(* IEC 61131-3 sources: Lasal-MCP/examples/SampleSource/2_PumpControlSolution/Stations/MachineControl/MachineControl/Class/SdiasSafetyManagerFSoE (part 2) *)

                          elsif (OptionalSettings.ModuleIDHBG = sHBG.usExpectedDeviceID) then
                            // the configured ID of LASAL and safety designer are equal

                            // if the module ID found is also the same => everthing is fine
                            if aModuleIDs[HBGPlace] = sHBG.usExpectedDeviceID then
                              MyPara.aPara[0] := _ClassOk$DINT;
                              CanActive := OldCanActive := TRUE;
                            else
                              // found something else
                              LogError("@02B4 (SdiasSafetyManagerFSoE::ClassSvr::NewInst) Wrong safety CAN terminal found (config of safety designer and hw classes match)");
                              MyPara.aPara[0] := _WrongHardware$DINT;
                              bHWConfigError := TRUE;
                            end_if;
                          else
                            // configuration of safety designer and hw classes does not match
                            LogError("@02B5 (SdiasSafetyManagerFSoE::ClassSvr::NewInst) Safety CAN terminal in hardware class configuration differs from safety designer configuration.");
                            MyPara.aPara[0] := _InvalidConfguration$DINT;
                            bHWConfigError := TRUE;
                          end_if;
                        else
                          MyPara.aPara[1] := SDIAS_SAFETY_INVALID_DEVICE_ID;

                          // projected in LASAL but not found in hardware
                          if sHBG.sdRequired then
                            MyPara.aPara[0] := _RequiredError$DINT;
                            bRequiredError := TRUE;
                            LogError("@02B6 (SdiasSafetyManagerFSoE::ClassSvr::NewInst) Required safety CAN terminal not available!");
                          else
                            // module is configured in safety designer
                            if (OptionalSettings.ModuleIDHBG <> SDIAS_SAFETY_INVALID_DEVICE_ID) then
                              // if the configuration does not match with the hardware classes
                              if (OptionalSettings.ModuleIDHBG <> sHBG.usExpectedDeviceID) then
                                LogError("@02B5 (SdiasSafetyManagerFSoE::ClassSvr::NewInst) Safety CAN terminal in hardware class configuration differs from safety designer configuration.");
                                MyPara.aPara[0] := _InvalidConfguration$DINT;
                                bHWConfigError := TRUE;

                              // the IDs match but it's not optional. since it's not available => error
                              elsif (OptionalSettings.OptionalFlagHBG.1 = FALSE) then
                                MyPara.aPara[0] := _NoHardware$DINT;
                                LogError("@02B7 (SdiasSafetyManagerFSoE::ClassSvr::NewInst) Could not find the non-optional Safety CAN terminal defined in the safety designer configuration.");
                                bHWConfigError := TRUE;

                              else
                                // if the IDs match and it's optional => just show no hardware (no error)
                                MyPara.aPara[0] := _NoHardware$DINT;
                              end_if;
                            else
                              LogError("@02B8 (SdiasSafetyManagerFSoE::ClassSvr::NewInst) Safety CAN terminal in hardware class configuration but not physically available and not in safety designer configuration.");
                              MyPara.aPara[0] := _NoHardware$DINT;
                            end_if;
                          end_if;
                        end_if;
                        sHBG.pThis^.NewInst(#MyPara, #MyResult);
                      else
                        // nothing projected for HBG in the lasal project

                        // if module is configured in safety designer
                        if (OptionalSettings.ModuleIDHBG <> SDIAS_SAFETY_INVALID_DEVICE_ID) then
                          // if a HBG has been found
                          if HBGPlace <> SDIAS_SAFETY_INVALID_MAX_PLACE then
                            // if it's not the configured module
                            if (aModuleIDs[HBGPlace] <> OptionalSettings.ModuleIDHBG) then
                              LogError("@02B9 (SdiasSafetyManagerFSoE::ClassSvr::NewInst) Safety CAN terminal found doesn't match the safety designer configuration.");
                              bHWConfigError := TRUE;
                            end_if;
                          else
                            // module not available (only a problem if it's not optional)
                            if (OptionalSettings.OptionalFlagHBG.1 = FALSE) then
                              LogError("@02BA (SdiasSafetyManagerFSoE::ClassSvr::NewInst) Could not find the non-optional Safety CAN terminal defined in the safety designer configuration.");
                              bHWConfigError := TRUE;
                            end_if;
                          end_if;
                        else
                          // module not configured in safety designer. if there is a module available, the number of IOs in safety does not match the config
                          if HBGPlace <> SDIAS_SAFETY_INVALID_MAX_PLACE then
                            LogError("@02BB (SdiasSafetyManagerFSoE::ClassSvr::NewInst) Safety CAN terminal found but not projected in the safety designer configuration.");
                            bHWConfigError := TRUE;
                          end_if;
                        end_if;
                      end_if;
                    else
                      // old firmware (no optional settings available)
                      if MaxPlace <> SDIAS_SAFETY_INVALID_MAX_PLACE then
                        pSafetyModuleInfo := #aSafetyModuleInfo[0];

                        // always the same command
                        MyPara.uiCmd := SDIAS_SET_CLASS_STATE;

                        for i := 0 to MaxPlace do
                          if pSafetyModuleInfo^.pThis then
                            MyPara.aPara[1] := aModuleIDs[i];
                            if aModuleIDs[i] = pSafetyModuleInfo^.usExpectedDeviceID then
                              MyPara.aPara[0] := _ClassOk$DINT;
                            elsif aModuleIDs[i] <> SDIAS_SAFETY_INVALID_DEVICE_ID then
                              if pSafetyModuleInfo^.sdRequired then
                                MyPara.aPara[0] := _RequiredError$DINT;
                                bRequiredError := TRUE;
                                LogValue("@02AC (SdiasSafetyManagerFSoE::ClassSvr::NewInst) Wrong safety IO module at required place {0}.", Value:=i);
                              else
                                MyPara.aPara[0] := _WrongHardware$DINT;
                                bHWConfigError  := TRUE;
                              end_if;
                            else
                              if pSafetyModuleInfo^.sdRequired then
                                MyPara.aPara[0] := _RequiredError$DINT;
                                bRequiredError := TRUE;
                                LogValue("@02AB (SdiasSafetyManagerFSoE::ClassSvr::NewInst) No safety IO module at required place {0}.", Value:=i);
                              else
                                MyPara.aPara[0] := _NoHardware$DINT;
                                // Hardwareclass placed in Project but no physical Hardware available is allowed
                                // bHWConfigError  := TRUE;
                              end_if;
                            end_if;
                            pSafetyModuleInfo^.pThis^.NewInst(#MyPara, #MyResult);

                          elsif aModuleIDs[i] <> SDIAS_SAFETY_INVALID_DEVICE_ID then  // HWK this pointer is NIL but a module is identified
                            bHWConfigError  := TRUE;
                          end_if;

                          pSafetyModuleInfo += sizeof(t_SdiasSafetyModuleInfo);
                        end_for;
                      end_if;

                      // Check if a module info was passed for which there is no corrosponding HWK object.
                      if MaxPlace + 1 < sizeof(t_ModuleIDs) then
                        // it's only a config error if it's not the HBG
                        if (aModuleIDs[MaxPlace + 1] <> SDIAS_SAFETY_INVALID_DEVICE_ID) & ((MaxPlace + 1) <> HBGPlace) then
                          bHWConfigError  := TRUE;
                        end_if;
                      end_if;

                      // check for hbg
                      if sHBG.pThis then
                        MyPara.uiCmd := SDIAS_SET_CLASS_STATE;
                        if HBGPlace <> SDIAS_SAFETY_INVALID_MAX_PLACE then
                          MyPara.aPara[1] := aModuleIDs[HBGPlace];

                          if aModuleIDs[HBGPlace] = sHBG.usExpectedDeviceID then
                            MyPara.aPara[0] := _ClassOk$DINT;
                            CanActive := OldCanActive := TRUE;
                            bHWConfigError := FALSE;
                          elsif aModuleIDs[HBGPlace] <> SDIAS_SAFETY_INVALID_DEVICE_ID then
                            if sHBG.sdRequired then
                              MyPara.aPara[0] := _RequiredError$DINT;
                              bRequiredError := TRUE;
                              LogError("@02BE (SdiasSafetyManagerFSoE::ClassSvr::NewInst) Wrong safety IO module at required HBG place.");
                            else
                              MyPara.aPara[0] := _WrongHardware$DINT;
                              CanActive := OldCanActive := FALSE;
                            end_if;
                          else
                            if sHBG.sdRequired then
                              MyPara.aPara[0] := _RequiredError$DINT;
                              bRequiredError := TRUE;
                              LogError("@02BF (SdiasSafetyManagerFSoE::ClassSvr::NewInst) HBG required but not available!");
                            else
                              MyPara.aPara[0] := _NoHardware$DINT;
                              CanActive := OldCanActive := FALSE;
                            end_if;
                          end_if;
                        else
                          MyPara.aPara[1] := SDIAS_SAFETY_INVALID_DEVICE_ID;
                          if sHBG.sdRequired then
                            MyPara.aPara[0] := _RequiredError$DINT;
                            bRequiredError := TRUE;
                            LogError("@02BE (SdiasSafetyManagerFSoE::ClassSvr::NewInst) Wrong safety IO module at required HBG place.");
                          else
                            MyPara.aPara[0] := _WrongHardware$DINT;
                            CanActive := OldCanActive := FALSE;
                          end_if;
                        end_if;
                        sHBG.pThis^.NewInst(#MyPara, #MyResult);
                      end_if;
                    end_if;

                    if bRequiredError then
                      MyPara.uiCmd := _BUS_IF_SET_REQUIRED_ERROR;
                      ToBusInterface.NewInst(#MyPara, #MyResult);
                    end_if;

                    if bHWConfigError then
                      // if we have optional settings, we already logged the reason
                      if b_GotOptionalSettings = FALSE then
                        LogError("@ß02C0 (SdiasSafetyManagerFSoE::ClassSvr::NewInst) Hardwareconfiguration does not match objects placed in network.");
                      end_if;

                      // Check if Safetymanyger is required
                      MyPara.uiCmd     := _BUS_IF_GET_REQUIRED_SETTING;
                      ToBusInterface.NewInst(pPara:=#MyPara, pResult:=#MyResult);
                      if MyResult.aData[0]$t_BusIFRetvalErrorcode = _BUS_IF_RETVAL_OK then
                        // if it's required => set required error
                        if MyResult.aData[4] then

                          MyPara.uiCmd := _BUS_IF_SET_REQUIRED_ERROR;
                          ToBusInterface.NewInst(#MyPara, #MyResult);
                        else

                          SetSafetyState(_WrongSafetyHW);
                          Online      := 0;

                          // Update BusIF ClassState
                          MyPara.uiCmd := _BUS_IF_SET_CLASS_STATE;
                          MyPara.aPara[0] := _WrongHardware$DINT;
                          ToBusInterface.NewInst(#MyPara, #MyResult);

                          // Cancel init
                          eInitSSWErrorStep := eInitSSW;
                          eInitSSW := _InitError;

                          // Set Module states
                          pSafetyModuleInfo := #aSafetyModuleInfo[0];
                          // always the same command
                          MyPara.uiCmd := SDIAS_SET_CLASS_STATE;
                          MyPara.aPara[0] := _ModuleFoundButManagerIsOff$DINT;

                          if MaxPlace <> SDIAS_SAFETY_INVALID_MAX_PLACE then
                            for i := 0 to MaxPlace do
                              if pSafetyModuleInfo^.pThis then
                                MyPara.aPara[1] := aModuleIDs[i];
                                pSafetyModuleInfo^.pThis^.NewInst(#MyPara, #MyResult);
                              end_if;
                              pSafetyModuleInfo += sizeof(t_SdiasSafetyModuleInfo);
                            end_for;
                          end_if;

                          // check for hbg
                          if sHBG.pThis then
                            sHBG.pThis^.NewInst(#MyPara, #MyResult);
                          end_if;

                        end_if;

                      end_if;

                    end_if;

                  else
                    LogError("@02C1 (SdiasSafetyManagerFSoE::ClassSvr::NewInst) Invalid SDO response buffer pointer.");
                  end_if;
                else
                  LogError("@02C2 (SdiasSafetyManagerFSoE::ClassSvr::NewInst) Invalid length for SDO response data.");
                end_if;

                eResponseState := _valid;
              else
                LogError("@02C3 (SdiasSafetyManagerFSoE::ClassSvr::NewInst) SDO response arrived when no response was expected.");
              end_if;
            end_if;
          elsif (LastSDO.Command = _BUS_IF_READ_VIA_SDO_CTRL) then
            if LastSDO.ResponseArrived = FALSE then
              if pPara^.aPara[5] = LastSDO.Length then
                if pPara^.aPara[4] then
                  // all parameters are fine, so we're ready
                  ret_code := READY;

                  // copy the response data
                  _memcpy(ptr1:=Config.pActData, ptr2:=pPara^.aPara[4]$pVoid, cntr:=LastSDO.Length);
                else
                  LogError("@02C1 (SdiasSafetyManagerFSoE::ClassState::NewInst) Invalid SDO response buffer pointer.");
                end_if;
              else
                LogError("@02C2 (SdiasSafetyManagerFSoE::ClassState::NewInst) Invalid length for SDO response data.");
              end_if;

              LastSDO.ResponseArrived := TRUE;
            else
              LogError("@02C3 (SdiasSafetyManagerFSoE::ClassState::NewInst) SDO response arrived when no response was expected.");
            end_if;
          elsif (LastSDO.Command = _BUS_IF_WRITE_VIA_SDO_CTRL) then
            if LastSDO.ResponseArrived = FALSE then
              // all parameters are fine, so we're ready
              ret_code := READY;

              LastSDO.ResponseArrived := TRUE;
            else
              LogError("@02C3 (SdiasSafetyManagerFSoE::ClassState::NewInst) SDO response arrived when no response was expected.");
            end_if;
          end_if;
        else
          LogError("@02C4 (SdiasSafetyManagerFSoE::ClassSvr::NewInst) SDO transfer failed.");
        end_if;
      else
        LogError("@02C5 (SdiasSafetyManagerFSoE::ClassSvr::NewInst) Received invalid SDO response.");
      end_if;

//**********************************************************************************************************************************************************
    _BUS_IF_DATA_POINTER_AVAILABLE:
      // does nothing in the FSoE version
      ret_code := READY;

//**********************************************************************************************************************************************************
    _BUS_IF_RESET_DETECTED:
      // don't overwrite other errors
      if SafetyState = _SafetyClassOK then
        SafetyState := _LostPowerSupply;
      end_if;

      // check if module is requred
      MyPara.uiCmd     := _BUS_IF_GET_REQUIRED_SETTING;
      ToBusInterface.NewInst(pPara:=#MyPara, pResult:=#MyResult);
      if MyResult.aData[0]$t_BusIFRetvalErrorcode = _BUS_IF_RETVAL_OK then
        // if it's required => set required error
        if MyResult.aData[4] then

          MyPara.uiCmd := _BUS_IF_SET_REQUIRED_ERROR;
          ToBusInterface.NewInst(#MyPara, #MyResult);
        end_if;
      end_if;

      // drop config of connected modules

      // initialize the message for the periphery
      MyPara.uiCmd := SDIAS_SET_CLASS_STATE;
      MyPara.aPara[1] := 0;// no device ID
      MyPara.aPara[0] := _NoHardware$DINT;

      // tell the connected IO module objects
      if MaxPlace <> SDIAS_SAFETY_INVALID_MAX_PLACE then
        pSafetyModuleInfo := #aSafetyModuleInfo[0];

        for i := 0 to MaxPlace do
          if pSafetyModuleInfo^.pThis then
            pSafetyModuleInfo^.pThis^.NewInst(#MyPara, #MyResult);
          end_if;

          pSafetyModuleInfo += sizeof(t_SdiasSafetyModuleInfo);
        end_for;
      end_if;

      // tell the hbg (if available)
      if sHBG.pThis then
        sHBG.pThis^.NewInst(#MyPara, #MyResult);
      end_if;

//**********************************************************************************************************************************************************
    _BUS_IF_RESET_GONE_DETECTED:
      if SafetyState = _LostPowerSupply then

        // get safety and serial numbers of connected modules
        bUpdateModuleConfig := TRUE;

        // remember the time. in case we don't get the SDO response to signal the firmware being ready, we use a timeout
        ud_ResetGoneTime := ops.tAbsolute;

        // we wait for an asynchronous SDO response in the cyclic of the base class. once we got that, the firmware is ready
        b_WaitForFirmwareBoot := TRUE;

        // refetch IDs of connected modules
        eCheckIDSSW := _Wait4Idle;

        SafetyState := _SafetyClassOK;
      end_if;

//**********************************************************************************************************************************************************

    CMD_GET_HARDWARE_DIAGNOSIS:
      //Returns module info
      ret_code := ERROR;
      pResult^.aData[0]$t_HWCGetHardwareDiagnosisOut.retcode := _HWC_RETVAL_ERROR;

      pStr_HWTRequested := pPara^.aPara[0]$t_HWCGetHardwareDiagnosisIn.pStr_HardewareTreeEntry;

      tmpplace := (pStr_HWTRequested+pPara^.aPara[0]$t_HWCGetHardwareDiagnosisIn.us_current_index)^$USINT;

      //Check if pointer is valid
      if aSafetyModuleInfo[tmpplace].pThis then

        // Set Offline Device ID
        pResult^.aData[0]$t_HWCGetHardwareDiagnosisOut.ud_DeviceID := (aSafetyModuleInfo[tmpplace].usExpectedDeviceID AND 2#00111000 ) shr 3;   // Bit 3-5 Modul typ
        pResult^.aData[0]$t_HWCGetHardwareDiagnosisOut.ud_Variante :=  aSafetyModuleInfo[tmpplace].usExpectedDeviceID AND 2#00000111;  // Bit 0-2 Submodul typ

        if aModuleIDs[tmpplace] = aSafetyModuleInfo[tmpplace].usExpectedDeviceID then

          ret_code := READY;
          pResult^.aData$t_HWCGetHardwareDiagnosisOut.retcode := _HWC_RETVAL_OK;

          pResult^.aData[0]$t_HWCGetHardwareDiagnosisOut.ud_DeviceID  := (aModuleIDs[tmpplace] AND 2#00111000 ) shr 3;  // Bit 3-5 Modul typ
          pResult^.aData[0]$t_HWCGetHardwareDiagnosisOut.ud_Variante  :=  aModuleIDs[tmpplace] AND 2#00000111; // // Bit 0-2 Submodul typ
          pResult^.aData[0]$t_HWCGetHardwareDiagnosisOut.ud_Place     := tmpplace;

          // Get Serialno ---------------------------------------------------------------------------------------------
          _memcpy(ptr1 := #a_SerialNo[0]
                , ptr2 := #sSafetySerNrs.aSerialNumbers[tmpplace]
                , cntr := sizeof(sSafetySerNrs.aSerialNumbers[tmpplace]) );

          a_SerialNo[sizeof(sSafetySerNrs.aSerialNumbers[tmpplace])] := 0;  // 0 Terminierung

          pResult^.aData[0]$t_HWCGetHardwareDiagnosisOut.pStr_SerialNo := #a_SerialNo[0];

          pResult^.aData[0]$t_HWCGetHardwareDiagnosisOut.hd_SafetyNumber  := sSafetySerNrs.aSafetyNumbers[tmpplace];

          // first free the old then create the memory (linked list) for the additional information

          if pAdditionalDiagInfo then
            HwDiagFreeDynExtList(pList:=pAdditionalDiagInfo);
          end_if;
          pAdditionalDiagInfo      := NIL;

          // add the firmware version
          pNewElement := HwDiagAddDynExt2List(ppList:=#pAdditionalDiagInfo, EntryID:=_HWC_DIAG_ID_SAFETY_FIRMWARE_VERSION, udVersion:=1, udDataLength:=sizeof(HDINT));

          if pNewElement then
            // add the data in the reserved memory
            (pNewElement$^HDINT + sizeof(t_HWCGetHardwareDiagnosisOutDynExt))^ := FirmwareVersion;
          end_if;

          // add the safety designer project name
          pNewElement := HwDiagAddDynExt2List(ppList:=#pAdditionalDiagInfo, EntryID:=_HWC_DIAG_ID_SAFETY_DESIGNER_PROJECT_NAME, udVersion:=1, udDataLength:=ProjectNameStr.GetLength());

          if pNewElement then
            // add the data in the reserved memory
            ProjectNameStr.ReadDataOff(udOff:=0, pData:=pNewElement$^USINT + sizeof(t_HWCGetHardwareDiagnosisOutDynExt), udMax:=pNewElement^.ud_DataLength);
          end_if;

          // add the safety designer project revision
          pNewElement := HwDiagAddDynExt2List(ppList:=#pAdditionalDiagInfo, EntryID:=_HWC_DIAG_ID_SAFETY_DESIGNER_PROJECT_REVISION, udVersion:=1, udDataLength:=ProjectRevisionStr.GetLength());

          if pNewElement then
            // add the data in the reserved memory
            ProjectRevisionStr.ReadDataOff(udOff:=0, pData:=pNewElement$^USINT + sizeof(t_HWCGetHardwareDiagnosisOutDynExt), udMax:=pNewElement^.ud_DataLength);
          end_if;

          pResult^.aData[0]$t_HWCGetHardwareDiagnosisOut.p_DynExtList := pAdditionalDiagInfo;

        elsif aModuleIDs[tmpplace] <> SDIAS_SAFETY_INVALID_DEVICE_ID then
          pResult^.aData$t_HWCGetHardwareDiagnosisOut.retcode := _HWC_RETVAL_ERROR_WRONG_HARDWARE;
        else
          pResult^.aData$t_HWCGetHardwareDiagnosisOut.retcode := _HWC_RETVAL_ERROR_NO_HARDWARE;
        end_if;

      else
        pResult^.aData[0]$t_HWCGetHardwareDiagnosisOut.retcode := _HWC_RETVAL_ERROR_SDIAS_MODULE_NOT_FOUND;
      end_if;

//**********************************************************************************************************************************************************
    CMD_GET_HARDWARE_TREE_ENTRY:
      //Returns module info

      ret_code := ERROR;
      pResult^.aData[0]$t_HWCGetHardwareTreeEntryOut.retcode := _HWC_RETVAL_ERROR;

      pStr_HWTreeEntry := pPara^.aPara[0]$t_HWCGetHardwareTreeEntryIn.pStr_LastHardewareTreeEntry;

      //First HWT Path
      if (pStr_HWTreeEntry + pStr_HWTreeEntry$^UINT^)^ <> HWT_ESCAPE_INTERNALBUS_SDIAS_SAFETY then  // + 1 for Byte length -1 for 2nd last element of string

        if aSafetyModuleInfo[0].pThis then

          _memcpy(ptr1 := #a_HWTEntryStr[0]
                , ptr2 := pPara^.aPara[0]$t_HWCGetHardwareTreeEntryIn.pStr_LastHardewareTreeEntry
                , cntr := pPara^.aPara[0]$t_HWCGetHardwareTreeEntryIn.pStr_LastHardewareTreeEntry$^UINT^ +2 );  // +2 2 Byte Strlength is not included in the stringlength

          // Add escape sequence
          a_HWTEntryStr[0]$UINT += 1;
          a_HWTEntryStr[a_HWTEntryStr[0]$UINT+1] := HWT_ESCAPE_INTERNALBUS_SDIAS_SAFETY;

          // Add Place
          a_HWTEntryStr[0]$UINT += 1;
          a_HWTEntryStr[a_HWTEntryStr[0]$UINT+1] := 0;

          //Return Hardware Tree Entry and set return codes
          pResult^.aData[0]$t_HWCGetHardwareTreeEntryOut.pStr_NextHardewareTreeEntry := #a_HWTEntryStr[0];

          pResult^.aData[0]$t_HWCGetHardwareTreeEntryOut.retcode := _HWC_RETVAL_OK_HWTSTR_RETURNED;
          ret_code := READY;

        else
          pResult^.aData[0]$t_HWCGetHardwareTreeEntryOut.retcode := _HWC_RETVAL_ERROR_SDIAS_MODULE_NOT_FOUND;
        end_if;

      //search next module
      else

        usNextPlace := (pStr_HWTreeEntry  + pPara^.aPara[0]$t_HWCGetHardwareTreeEntryIn.us_current_index)^$USINT+1;

        if usNextPlace <= SDIAS_SAFETY_MAX_PLACE_NR &
           aSafetyModuleInfo[usNextPlace].pThis then

          _memcpy(ptr1 := #a_HWTEntryStr[0]
                , ptr2 := pPara^.aPara[0]$t_HWCGetHardwareTreeEntryIn.pStr_LastHardewareTreeEntry
                , cntr := pPara^.aPara[0]$t_HWCGetHardwareTreeEntryIn.pStr_LastHardewareTreeEntry$^UINT^ +2 );  // +2 2 Byte Strlength is not included in the stringlength

          // Set new Place
          a_HWTEntryStr[a_HWTEntryStr[0]$UINT + 1] := usNextPlace;

          pResult^.aData[0]$t_HWCGetHardwareTreeEntryOut.pStr_NextHardewareTreeEntry := #a_HWTEntryStr[0];

          //Return Hardware Tree Entry and set return codes
          pResult^.aData[0]$t_HWCGetHardwareTreeEntryOut.retcode := _HWC_RETVAL_OK_HWTSTR_RETURNED;
          ret_code := READY;

        else
          ret_code := READY;
          pResult^.aData$t_HWCGetHardwareTreeEntryOut.retcode := _HWC_RETVAL_OK_END_OF_LIST;
        end_if;
      end_if;

//**********************************************************************************************************************************************************

//*****************************************************************************
//** INTERNAL COMMANDS                                                       **
//*****************************************************************************

//**********************************************************************************************************************************************************
    CMD_SM_READ_PDO_SIZE:
      // get the size of the PDO
      LastSDO.Command := _BUS_IF_READ_VIA_SDO;
      LastSDO.Offset  := SBF_OFFSET_SPDO_LENGTH;
      LastSDO.Length  := sizeof(UINT);

      MyPara.uiCmd    := LastSDO.Command$UINT;
      MyPara.aPara[0] := LastSDO.Offset;
      MyPara.aPara[1] := LastSDO.Length;
      ret_code := ToBusInterface.NewInst(#MyPara, #MyResult);

//**********************************************************************************************************************************************************
  else
    ret_code := SafetyBaseFSoE::NewInst(pPara, pResult);
//**********************************************************************************************************************************************************
  END_CASE;

END_FUNCTION

FUNCTION VIRTUAL SdiasSafetyManagerFSoE::ShowProjectRevision

  ProjectNameStr.WriteDataOff(udLen:=PrjNameStrLen + 1, udOff:=0, pData:=pPrjNameStr);

  ProjectRevisionStr.WriteDataOff(udLen:=PrjRevStrLen + 1, udOff:=0, pData:=pPrjRevStr);

END_FUNCTION

FUNCTION VIRTUAL SdiasSafetyManagerFSoE::InitSafeModule
  VAR_OUTPUT
    sd_retval 	: DINT;
  END_VAR

  // allocate memory for finding unsafe-IO-Servers
  // in first place we allocate 512 byte for our blocked transfers
  p_BlockedTransferMemory := ToStdLib.Malloc( size := SBF_CONFIG_MEMORY_BLOCK_SIZE );
  IF p_BlockedTransferMemory <> NIL THEN
    ud_BlockedTransferMemorySize := SBF_CONFIG_MEMORY_BLOCK_SIZE;
  ELSE
    SafetyState := _MemAllocFailed;
    sd_retval := -100;
    return;
  END_IF;

  // if there is a safety manager to gather the configuration
  if pSafetyManagerThis then
    // allocate memory for gathering configuration information => in first place we allocate 512 byte
    pConfigMem := ToStdLib.Malloc( size := SBF_CONFIG_MEMORY_BLOCK_SIZE );
    IF pConfigMem <> NIL THEN
      ConfigMemSize := SBF_CONFIG_MEMORY_BLOCK_SIZE;
      ConfigMemSizeUsed := 4;
    ELSE
      SafetyState := _MemAllocFailed;
      sd_retval := -100;
      return;
    END_IF;
  end_if;

END_FUNCTION

FUNCTION VIRTUAL GLOBAL SdiasSafetyManagerFSoE::CanOut::NewInst
  VAR_INPUT
    pPara 	: ^CmdStruct;
    pResult 	: ^results;
  END_VAR
  VAR_OUTPUT
    ret_code 	: iprStates;
  END_VAR
  VAR
    tempCmd         : CmdStruct;
    _result         : results;
  END_VAR

  CASE pPara^.uiCmd OF
//**********************************************************************************************************************************************************
    SDIAS_SAFETY_LOGIN_HBG:
      // check parameters
      if pPara^.aPara[0] & pPara^.aPara[1] then

        sHBG.pThis               := pPara^.aPara[0]$pVirtualBase;
        sHBG.usExpectedDeviceID  := pPara^.aPara[1]$USINT;
        sHBG.sdRequired          := pPara^.aPara[2];
        sHBG.pIOStates           := pPara^.aPara[3]$^HDINT;

        // if leds/hgb not added so far, add them
        if StateBytesUsed = 0 then
          StateBitsUsed := (sizeof(t_LedAndIOStates.biLEDs) + sizeof(t_LedAndIOStates.HBGInputs)) * 8;
          // refresh state bytes used value
          StateBytesUsed := ((StateBitsUsed-1) / 8) + 1;
        end_if;

        if sHBG.sdRequired & (b_AnyModuleRequired = FALSE) then
          b_AnyModuleRequired := TRUE;
          // if any access is required => the businterface is also required
          tempCmd.uiCmd := _BUS_IF_SET_REQUIRED;
          ToBusInterface.NewInst(pPara:=#tempCmd, pResult:=#_result);
          if _result.aData[0]$t_BusIFRetvalErrorcode <> _BUS_IF_RETVAL_OK then
            LogError("@029D (SdiasSafetyManagerFSoE::CanOut::NewInst) Failed to set the BusInterface to required.");
          end_if;
        end_if;
      else
        ret_code := ERROR;
      end_if;
//**********************************************************************************************************************************************************
  END_CASE;

  ret_code := READY;

END_FUNCTION

FUNCTION VIRTUAL SdiasSafetyManagerFSoE::GetConfiguration
  VAR
    pHelp                 : ^void;
    SizeToGo              : UINT;
    ActSize               : UINT;
    ActAddr               : HDINT;
    SDOReqBuf             : SDORequReadConfig;
    SDORspBuf             : ARRAY [0..SBF_SDO_MAX_LENGTH-1] OF USINT;
    pRspBuf               : ^SDORespReadConfig;
    i                     : DINT;
    pSafetyModuleInfo     : ^t_SdiasSafetyModuleInfo;
    MyPara 	              : CmdStruct;
    MyResult              : Results;
  END_VAR

  //initialize header-data for request

  //calculate length without crc
  SDOReqBuf.StdHeader.Len := sizeof(SDORequReadConfig) - sizeof(SDOHeader.StdHeader.CRC);

  //type
  SDOReqBuf.StdHeader.Typ := SDO_STD;

  //command for reading config data
  SDOReqBuf.StdHeader.Cmd := SBF_SDO_COMMAND_READ;

  // read the complete 256 Bytes of safety and serial number info
  pHelp    := #sSafetySerNrs;
  SizeToGo := sizeof(sSafetySerNrs);
  pRspBuf  := (#SDORspBuf)$^SDORespReadConfig;
  ActAddr  := SBF_SDO_ADDRESS_SER_NR_DATA;

  while SizeToGo do
    if SizeToGo > SDIAS_SAFTEY_SDO_MAX_DATA_PER_PAKET then
      ActSize := SDIAS_SAFTEY_SDO_MAX_DATA_PER_PAKET;
    else
      ActSize := SizeToGo;
    end_if;

    if SDOReadCfgRequ(p_SDORequestBuffer  := #SDOReqBuf,
                      p_SDOResponseBuffer := pRspBuf,
                      ud_Address          := ActAddr,
                      us_Length           := ActSize$USINT,
                      b_UseCache          := FALSE) then
      LogError("@02C6 (SdiasSafetyManagerFSoE::GetConfiguration) Failed to get safety and serial numbers of the IO modules.");
      return;
    else
      _memcpy(ptr1:=pHelp, ptr2:=#pRspBuf^.ud_Data, cntr:=ActSize);
    end_if;

    SizeToGo  -= ActSize;
    ActAddr   += ActSize;
    pHelp     += ActSize;
  end_while;

  // read the complete 64 Bytes of hardware version info
  pHelp    := #sHwVersions;
  SizeToGo := sizeof(sHwVersions);
  pRspBuf  := (#SDORspBuf)$^SDORespReadConfig;
  ActAddr  := SBF_SDO_ADDRESS_HW_VERSIONS;

  while SizeToGo do
    if SizeToGo > SDIAS_SAFTEY_SDO_MAX_DATA_PER_PAKET then
      ActSize := SDIAS_SAFTEY_SDO_MAX_DATA_PER_PAKET;
    else
      ActSize := SizeToGo;
    end_if;

    if SDOReadCfgRequ(p_SDORequestBuffer  := #SDOReqBuf,
                      p_SDOResponseBuffer := pRspBuf,
                      ud_Address          := ActAddr,
                      us_Length           := ActSize$USINT,
                      b_UseCache          := FALSE) then
      LogError("@02F9 (SdiasSafetyManagerFSoE::GetConfiguration) Failed to get hw versions of the Safe IO modules!");
      return;
    else
      // if the return code in the response buffer is not 0 => the virtual memory is not available
      if pRspBuf^.us_Returncode <> 0 then
        // reset array to make sure there are no hw versions stored
        _memset(dest:=#sHwVersions.aVersion[0], usByte:=0, cntr:=sizeof(sHwVersions));
        exit;
      end_if;

      _memcpy(ptr1:=pHelp, ptr2:=#pRspBuf^.ud_Data, cntr:=ActSize);
    end_if;

    SizeToGo  -= ActSize;
    ActAddr   += ActSize;
    pHelp     += ActSize;
  end_while;

  // only available for IOs, not the HBG
  if MaxPlace <> SDIAS_SAFETY_INVALID_MAX_PLACE then
    // always the same command
    MyPara.uiCmd := SDIAS_SET_NUMBERS;

    pSafetyModuleInfo := #aSafetyModuleInfo[0];
    for i := 0 to MaxPlace$DINT do
      // safety number
      MyPara.aPara[0] := (sSafetySerNrs.aSafetyNumbers[i])$DINT;

      // pointer to serial number string
      MyPara.aPara[1] := (#sSafetySerNrs.aSerialNumbers[i][0])$DINT;

      // hw version
      MyPara.aPara[2] := (sHwVersions.aVersion[i])$DINT;

      pSafetyModuleInfo^.pThis^.NewInst(#MyPara, #MyResult);

      pSafetyModuleInfo += sizeof(t_SdiasSafetyModuleInfo);
    end_for;
  end_if;

END_FUNCTION

FUNCTION VIRTUAL GLOBAL SdiasSafetyManagerFSoE::DisconnectEvent
  VAR
    i                 : UDINT;
    pSafetyModuleInfo : ^t_SdiasSafetyModuleInfo;
    MyPara 	          : CmdStruct;
    MyResult          : Results;
  END_VAR

  SafetyBaseFSoE::DisconnectEvent();

  // initialize the message for the periphery
  MyPara.uiCmd := SDIAS_SET_CLASS_STATE;
  MyPara.aPara[1] := 0;// no device ID
  MyPara.aPara[0] := _NoHardware$DINT;

  // tell the connected IO module objects
  if MaxPlace <> SDIAS_SAFETY_INVALID_MAX_PLACE then
    pSafetyModuleInfo := #aSafetyModuleInfo[0];

    for i := 0 to MaxPlace do
      if pSafetyModuleInfo^.pThis then
        pSafetyModuleInfo^.pThis^.NewInst(#MyPara, #MyResult);
      end_if;

      pSafetyModuleInfo += sizeof(t_SdiasSafetyModuleInfo);
    end_for;
  end_if;

  // tell the hbg (if available)
  if sHBG.pThis then
    sHBG.pThis^.NewInst(#MyPara, #MyResult);
  end_if;

  // clear the strings
  ProjectNameStr.Clear();
  ProjectRevisionStr.Clear();

END_FUNCTION

FUNCTION VIRTUAL SdiasSafetyManagerFSoE::SetSafetyState
  VAR_INPUT
    NewState 	: SafetyConfigStateType;
  END_VAR
  VAR
    MyPara 	  : CmdStruct;
    MyResult	: results;
  END_VAR

  // use it locally
  SafetyState := NewState;

  // tell the outer class
  MyPara.uiCmd := SDIAS_SET_SAFETY_STATE;
  MyPara.aPara[0] := NewState$DINT;
  ToBusInterface.NewInst(#MyPara, #MyResult);

END_FUNCTION

FUNCTION VIRTUAL GLOBAL SdiasSafetyManagerFSoE::CyWork
  VAR_INPUT
    EAX 	: UDINT;
  END_VAR
  VAR_OUTPUT
    state (EAX) 	: UDINT;
  END_VAR
  VAR
    MyPara 	          : CmdStruct;
    MyResult          : Results;
    TmpRetCode        : iprStates;
  END_VAR

  // if the initialisiation has been finished and there is an object for the hbg check if it's has been connected or disconnected
  if Online then

    case eCheckIDSSW of
  //**********************************************************************************************************************************************************
      _Nothing:
        if sHBG.pThis then
          // check for a can connect event
          if CanActive > OldCanActive then
            // if we're already idle => get it on
            if eResponseState = _idle then
              eCheckIDSSW := _GetIDs;
            else
              // otherwise, wait for it (need to remember the connect event)
              eCheckIDSSW := _Wait4Idle;
            end_if;

          // check for a can disconnect event
          elsif CanActive < OldCanActive then
            if sHBG.sdRequired then
              // if it's required => required error
              MyPara.uiCmd := _BUS_IF_SET_REQUIRED_ERROR;
              ToBusInterface.NewInst(#MyPara, #MyResult);
            else
              // otherwise show that it has been disconnected
              MyPara.uiCmd := SDIAS_SET_CLASS_STATE;
              MyPara.aPara[1] := 0;// no device ID
              MyPara.aPara[0] := _NoHardware$DINT;
              sHBG.pThis^.NewInst(#MyPara, #MyResult);
            end_if;
          end_if;
          OldCanActive := CanActive;
        end_if;

  //**********************************************************************************************************************************************************
      _Wait4Idle:
        if eResponseState = _idle then
          eCheckIDSSW := _GetIDs;
        end_if;

  //**********************************************************************************************************************************************************
      _GetIDs:
        case eResponseState of
        //*****************************************************
          _idle:
            LastSDO.Command := _BUS_IF_READ_VIA_SDO;
            LastSDO.Offset  := SBF_OFFSET_IO_MODULE_IDS;
            LastSDO.Length  := sizeof(t_ModuleIDs);

            MyPara.uiCmd    := LastSDO.Command$UINT;
            MyPara.aPara[0] := LastSDO.Offset;
            MyPara.aPara[1] := LastSDO.Length;
            TmpRetcode := ToBusInterface.NewInst(#MyPara, #MyResult);
            if TmpRetcode = READY then
              SDOTimeMark  := ops.tAbsolute;
              eResponseState:= _wait;
            elsif TmpRetcode = ERROR then
              LogError("@02A7 (SdiasSafetyManagerFSoE::InitModule) Failed to add read SDO for module configuration.");
            end_if;
        //*****************************************************
          _wait:
            // wait for response
            if ((ops.tAbsolute - SDOTimeMark) > SDIAS_SAFTEY_SDO_RESPONSE_TIMEOUT) then
              LogError("@02A1 (SdiasSafetyManagerFSoE::InitModule) SDO Response timeout while waiting for the module configuration.");
              eCheckIDSSW := _Nothing;
              eResponseState := _idle;
            end_if;
        //*****************************************************
          _valid:
            eCheckIDSSW := _Nothing;
            eResponseState := _idle;
        //*****************************************************
        end_case;
  //**********************************************************************************************************************************************************
    end_case;
  end_if;

  state := SafetyBaseFSoE::CyWork(0);

END_FUNCTION

FUNCTION VIRTUAL SdiasSafetyManagerFSoE::RefreshAsySrv
  VAR
    i                 : UDINT;
    pSafetyModuleInfo : ^t_SdiasSafetyModuleInfo;
    MyPara 	          : CmdStruct;
    MyResult          : Results;
    AsyValues         : t_AsyRefresh;
  END_VAR

  // tell the outer class
  MyPara.uiCmd := SDIAS_SET_ASY_STATE;
  AsyValues.QuitComError := QuitComError;
  MyPara.aPara[0] := (#AsyValues)$DINT;
  ToBusInterface.NewInst(#MyPara, #MyResult);

  // tell the connected IO module objects
  if MaxPlace <> SDIAS_SAFETY_INVALID_MAX_PLACE then
    pSafetyModuleInfo := #aSafetyModuleInfo[0];

    for i := 0 to MaxPlace do
      if pSafetyModuleInfo^.pThis then
        pSafetyModuleInfo^.pThis^.NewInst(#MyPara, #MyResult);
      end_if;

      pSafetyModuleInfo += sizeof(t_SdiasSafetyModuleInfo);
    end_for;
  end_if;

END_FUNCTION

FUNCTION VIRTUAL GLOBAL SdiasSafetyManagerFSoE::FastUnsafeOutputs::Write
  VAR_INPUT
    input (EAX) 	: BDINT;
  END_VAR
  VAR_OUTPUT
    result (EAX) 	: BDINT;
  END_VAR
  VAR
    pUnsafeOutLogin : ^t_FastUnsafeOuts;
  END_VAR

  // if the pointer is valid and we're in the first init run (the firstscan check prevents a crash caused by someone writing on the server during runtime)
  if input & (us_FirstScan < 2) then
    pUnsafeOutLogin := input$^t_FastUnsafeOuts;
    // check if it's the correct usage of the class
    if pUnsafeOutLogin^.Kennung = SDIAS_SAFETY_FAST_UNSAFE_KENNUNG then
      pFastUnsafeOutThis := pUnsafeOutLogin^.pThis;
    end_if;
  end_if;

  result := input;

END_FUNCTION

FUNCTION VIRTUAL GLOBAL SdiasSafetyManagerFSoE::FastUnsafeInputs::Write
  VAR_INPUT
    input (EAX) 	: BDINT;
  END_VAR
  VAR_OUTPUT
    result (EAX) 	: BDINT;
  END_VAR

  FastUnsafeInputs := input;
  result := FastUnsafeInputs;

END_FUNCTION

FUNCTION VIRTUAL SdiasSafetyManagerFSoE::SetRetryCounter
  VAR
    pSafetyModuleInfo : ^t_SdiasSafetyModuleInfo;
    MyPara 	 : CmdStruct;
    MyResult : Results;
    i        :  USINT;
  END_VAR

  if b_RetryCounterAvailable then

    if MaxPlace <> SDIAS_SAFETY_INVALID_MAX_PLACE then
      //Command for new inst call in sdiassafetybase
      MyPara.uiCmd := SDIAS_SET_RETRY_COUNTER;

      //calls newinst method of all safety modules which exists.
      for i := 0 to MaxPlace do
        pSafetyModuleInfo := #aSafetyModuleInfo[i];
        MyPara.aPara[0] := a_RetryCnt[i];
        MyPara.aPara[1] := a_RetryCnt[i+16];  //+16 for retry counter of µC2
        pSafetyModuleInfo^.pThis^.NewInst(#MyPara, #MyResult);
      end_for;
    end_if;
  else
    //Retrycounter not available -> show -1 at servers.
    SafetyRetryCounter := -1; //Not available

    if MaxPlace <> SDIAS_SAFETY_INVALID_MAX_PLACE then
      MyPara.uiCmd := SDIAS_RETRY_COUNTER_NOT_AVAILABLE;
      for i := 0 to MaxPlace do
        pSafetyModuleInfo := #aSafetyModuleInfo[i];
        pSafetyModuleInfo^.pThis^.NewInst(#MyPara, #MyResult);
      end_for;
    end_if;
  end_if;

END_FUNCTION

FUNCTION VIRTUAL GLOBAL SdiasSafetyManagerFSoE::Background
  VAR_INPUT
    EAX 	: UDINT;
  END_VAR
  VAR_OUTPUT
    state (EAX) 	: UDINT;
  END_VAR

  // if we have to update the module config, are not busy and the firmware has already booted (or a timeout on the boot occured)
  if bUpdateModuleConfig & (eCheckIDSSW = _Nothing) & ((b_WaitForFirmwareBoot = FALSE) | ((ops.tAbsolute - ud_ResetGoneTime) > SBF_FIRMWARE_BOOTUP_TIMEOUT)) then
    bUpdateModuleConfig := FALSE;

    GetConfiguration();
  end_if;

  state := SafetyBaseFSoE::Background(0);

END_FUNCTION

FUNCTION VIRTUAL SdiasSafetyManagerFSoE::BusConfigWrite
  VAR_INPUT
    Offset 	: HDINT;
    Length 	: UINT;
    pData 	: pVoid;
    IsControlAccess 	: BOOL;(* := FALSE *)
  END_VAR
  VAR_OUTPUT
    retcode 	: iprStates;
  END_VAR
  VAR
    TmpRetcode  : iprStates;
    MyPara      : CmdStruct;
    MyResult    : results;
  END_VAR

  retcode := BUSY;

  case Config.BusConfigSSW of
//**********************************************************************************************************************************************************
    _PrepareAccess:
      Config.RestLength := Length;
      Config.pActData   := pData;

      Config.BusConfigSSW := _StartAccess;

//**********************************************************************************************************************************************************
    _StartAccess:
      if IsControlAccess then
        LastSDO.Command := _BUS_IF_WRITE_VIA_SDO_CTRL;
      else
        LastSDO.Command := _BUS_IF_WRITE_VIA_SDO;
      end_if;

      LastSDO.Offset  := Offset$DINT;
      if Config.RestLength > SDIAS_SAFETY_MAX_SDO_DATA_PER_CYCLE then
        LastSDO.Length  := SDIAS_SAFETY_MAX_SDO_DATA_PER_CYCLE;
      else
        LastSDO.Length  := Config.RestLength;
      end_if;
      LastSDO.ResponseArrived := FALSE;

      MyPara.uiCmd    := LastSDO.Command;
      MyPara.aPara[0] := LastSDO.Offset;
      MyPara.aPara[1] := LastSDO.Length;
      MyPara.aPara[2] := Config.pActData$DINT;
      TmpRetcode := ToBusInterface.NewInst(#MyPara, #MyResult);
      if TmpRetcode = READY then
        Config.SDOTimeMark  := ops.tAbsolute;
        Config.BusConfigSSW := _Wait4Answer;
      elsif TmpRetcode = ERROR then
        retcode := ERROR;
        LogError("@02BC (SdiasSafetyManagerFSoE::BusConfigWrite) Failed to add write SDO for module configuration.");
      end_if;

//**********************************************************************************************************************************************************
    _Wait4Answer:
      // wait for response

      // check for response
      if LastSDO.ResponseArrived then
        Config.RestLength -= LastSDO.Length;
        Config.pActData   += LastSDO.Length;

        if Config.RestLength = 0 then
          retcode := READY;
          Config.BusConfigSSW := _PrepareAccess;
        end_if;
      elsif ((ops.tAbsolute - Config.SDOTimeMark) > SDIAS_SAFTEY_SDO_RESPONSE_TIMEOUT) then
        LogError("@02BD (SdiasSafetyManagerFSoE::BusConfigWrite) SDO Response timeout while waiting for the write response.");
        retcode := ERROR;
      end_if;

//**********************************************************************************************************************************************************
  end_case;

END_FUNCTION

FUNCTION VIRTUAL SdiasSafetyManagerFSoE::BusConfigRead
  VAR_INPUT
    Offset 	: HDINT;
    Length 	: UINT;
    pData 	: pVoid;
    IsControlAccess 	: BOOL;(* := FALSE *)
  END_VAR
  VAR_OUTPUT
    retcode 	: iprStates;
  END_VAR
  VAR
    TmpRetcode  : iprStates;
    MyPara      : CmdStruct;
    MyResult    : results;
  END_VAR

  retcode := BUSY;

  case Config.BusConfigSSW of
//**********************************************************************************************************************************************************
    _PrepareAccess:
      Config.RestLength := Length;
      Config.pActData   := pData;

      Config.BusConfigSSW := _StartAccess;

//**********************************************************************************************************************************************************
    _StartAccess:
      if IsControlAccess then
        LastSDO.Command := _BUS_IF_READ_VIA_SDO_CTRL;
      else
        LastSDO.Command := _BUS_IF_READ_VIA_SDO;
      end_if;

      LastSDO.Offset  := Offset$DINT;
      if Config.RestLength > SDIAS_SAFETY_MAX_SDO_DATA_PER_CYCLE then
        LastSDO.Length  := SDIAS_SAFETY_MAX_SDO_DATA_PER_CYCLE;
      else
        LastSDO.Length  := Config.RestLength;
      end_if;
      LastSDO.ResponseArrived := FALSE;

      MyPara.uiCmd    := LastSDO.Command;
      MyPara.aPara[0] := LastSDO.Offset;
      MyPara.aPara[1] := LastSDO.Length;
      TmpRetcode := ToBusInterface.NewInst(#MyPara, #MyResult);
      if TmpRetcode = READY then
        Config.SDOTimeMark  := ops.tAbsolute;
        Config.BusConfigSSW := _Wait4Answer;
      elsif TmpRetcode = ERROR then
        retcode := ERROR;
        LogError("@02BC (SdiasSafetyManagerFSoE::BusConfigRead) Failed to add write SDO for module configuration.");
      end_if;

//**********************************************************************************************************************************************************
    _Wait4Answer:
      // wait for response

      // check for response
      if LastSDO.ResponseArrived then
        Config.RestLength -= LastSDO.Length;
        Config.pActData   += LastSDO.Length;

        if Config.RestLength = 0 then
          retcode := READY;
          Config.BusConfigSSW := _PrepareAccess;
        end_if;
      elsif ((ops.tAbsolute - Config.SDOTimeMark) > SDIAS_SAFTEY_SDO_RESPONSE_TIMEOUT) then
        LogError("@02BD (SdiasSafetyManagerFSoE::BusConfigRead) SDO Response timeout while waiting for the write response.");
        retcode := ERROR;
      end_if;

//**********************************************************************************************************************************************************
  end_case;

END_FUNCTION

FUNCTION SdiasSafetyManagerFSoE::HwDiagFreeDynExtList
  VAR_INPUT
    pList 	: ^t_HWCGetHardwareDiagnosisOutDynExt;
  END_VAR
  VAR
    pHelp 	: ^t_HWCGetHardwareDiagnosisOutDynExt;
  END_VAR

  while pList do
    // remember the current entry
    pHelp := pList;

    // set plist to the next entry and free pHelp
    pList := pList^.p_Next;

    // free the current entry
    ToStdLib.Free(mptr:=pHelp);
  end_while;

END_FUNCTION

FUNCTION SdiasSafetyManagerFSoE::HwDiagAddDynExt2List
  VAR_INPUT
    ppList 	: ^t_pHWCGetHardwareDiagnosisOutDynExt;
    EntryID 	: t_HWCGetHardwareDiagnosisOutType;
    udVersion 	: UDINT;
    udDataLength 	: UDINT;
  END_VAR
  VAR_OUTPUT
    pNewElement 	: t_pHWCGetHardwareDiagnosisOutDynExt;
  END_VAR

  if ppList^ = NIL then
    ppList^$pVoid := ToStdLib.Malloc(size:=sizeof(t_HWCGetHardwareDiagnosisOutDynExt) + udDataLength);
    pNewElement := ppList^;
  else
    pNewElement := ppList^;
    while pNewElement^.p_Next <> NIL do
      pNewElement := pNewElement^.p_Next;
    end_while;
    pNewElement^.p_Next$pVoid := ToStdLib.Malloc(size:=sizeof(t_HWCGetHardwareDiagnosisOutDynExt) + udDataLength);
    pNewElement := pNewElement^.p_Next;
  end_if;

  if pNewElement <> NIL then
    // initialize the new memory
    pNewElement^.DiagID         := EntryID;
    pNewElement^.ud_Version     := udVersion;
    pNewElement^.p_Next         := NIL;
    pNewElement^.ud_DataLength  := udDataLength;

    if udDataLength then
      _memset(dest:=pNewElement + sizeof(t_HWCGetHardwareDiagnosisOutDynExt), usByte:=0, cntr:=udDataLength);
    end_if;
  end_if;

END_FUNCTION

FUNCTION VIRTUAL GLOBAL SdiasSafetyManagerFSoE::HGWOut::NewInst
  VAR_INPUT
    pPara 	: ^CmdStruct;
    pResult 	: ^Results;
  END_VAR
  VAR_OUTPUT
    ret_code 	: iprStates;
  END_VAR
  VAR
    tempCmd         : CmdStruct;
    _result         : results;
    dRetCode        : DINT;
    tempHWPath      : PathInfoType;
  END_VAR

  ret_code := READY;

  case pPara^.uiCmd of

    //**********************************************************************************************************************************************************
    SDIAS_SAFETY_GET_HGW_INFO:

      //Check for valid version
      //*****************************************************************************
      if pPara^.aPara[0] = 0x1 then

        //Return version number
        pResult^.aData[0] := 0x1;

        //pointer to input data to scp
        sHGW.pInputPDO           := pPara^.aPara[1]$^void;

        if sHGW.pInputPDO = nil then
          ret_code := ERROR;
          LogError(e_msg:="@03DD (SdiasSafetyManagerFSoE::HGWOut::NewInst) Pointer to input data of SCP is invalid.");
          return;
        end_if;

        // add PDO input data
        dRetCode :=  AddPDOToInputBuffer(ud_p2Buffer        := sHGW.pInputPDO$UDINT
                                      , ud_SafetyNr         := sHGW.hdSafetyNrb$UDINT
                                      , b_IsOptional        := FALSE
                                      , ui_PdoLen           := sHGW.InputPDOLength
                                      , ui_TargetOffset     := sHGW.InputPDOOffset
                                      );

        // return the pointer to the Buffer (is linear local memory, so the offset can be added later)
        sHGW.pOutputPDO$UDINT := GetPointer2PDOBuffer();

        pResult^.uiLng := 27;
        pResult^.aData[1]$UDINT := (sHGW.pOutputPDO+sHGW.OutputPDOOffset)$UDINT;
        pResult^.aData[5]$UINT  := sHGW.InputPDOLength;  //data to scp
        pResult^.aData[7]$UINT  := sHGW.OutputPDOLength; //data to hgw
        pResult^.aData[9]$UINT  := sHGW.uiSlotID;
        pResult^.aData[11]$UINT  := sHGW.uiCommunicationID;
        pResult^.aData[13]$USINT := sHGW.udMachineNrb$USINT;    //Old version, 1 byte machine number
        pResult^.aData[17]$USINT := sCPUConfig.CompPathLen$USINT;
        pResult^.aData[18]$UDINT := sCPUConfig.pCompPath$UDINT;
        pResult^.aData[22]$UDINT := sCPUConfig.SafetyNbr$UDINT;
        pResult^.aData[26]$UDINT := (#ErrorState)$UDINT;

      //Check for valid version
      //*****************************************************************************
      elsif pPara^.aPara[0] = 0x2 then

        //Return version number
        pResult^.aData[0] := 0x2;

        //pointer to input data to scp
        sHGW.pInputPDO           := pPara^.aPara[1]$^void;

        if sHGW.pInputPDO = nil then
          ret_code := ERROR;
          LogError(e_msg:="@03DD (SdiasSafetyManagerFSoE::HGWOut::NewInst) Pointer to input data of SCP is invalid.");
          return;
        end_if;

        // add PDO input data
        dRetCode :=  AddPDOToInputBuffer(ud_p2Buffer         := sHGW.pInputPDO$UDINT
                                      , ud_SafetyNr         := sHGW.hdSafetyNrb$UDINT
                                      , b_IsOptional        := FALSE
                                      , ui_PdoLen           := sHGW.InputPDOLength
                                      , ui_TargetOffset     := sHGW.InputPDOOffset
                                      );

        // return the pointer to the Buffer (is linear local memory, so the offset can be added later)
        sHGW.pOutputPDO$UDINT := GetPointer2PDOBuffer();

        pResult^.uiLng := 30;
        pResult^.aData[1]$UDINT := (sHGW.pOutputPDO+sHGW.OutputPDOOffset)$UDINT;
        pResult^.aData[5]$UINT  := sHGW.InputPDOLength;  //data to scp
        pResult^.aData[7]$UINT  := sHGW.OutputPDOLength; //data to hgw
        pResult^.aData[9]$UINT  := sHGW.uiSlotID;
        pResult^.aData[11]$UINT  := sHGW.uiCommunicationID;
        pResult^.aData[13]$UDINT := sHGW.udMachineNrb;
        pResult^.aData[17]$USINT := sCPUConfig.CompPathLen$USINT;
        pResult^.aData[18]$UDINT := sCPUConfig.pCompPath$UDINT;
        pResult^.aData[22]$UDINT := sCPUConfig.SafetyNbr$UDINT;
        pResult^.aData[26]$UDINT := (#ErrorState)$UDINT;

      //*****************************************************************************
      else
        // unknown version of the request
        ret_code := ERROR;
      end_if;

    //**********************************************************************************************************************************************************
    SDIAS_SAFETY_LOGIN_HGW:

      //Check for valid version
      if pPara^.aPara[0] = 0x1 then

      // check parameters
        if pPara^.aPara[1] then
          sHGW.pThis         := pPara^.aPara[1]$pVirtualBase; //this pointer of connect hgw communication class
          sHGW.sdRequired    := pPara^.aPara[2];              //required

        if sHGW.sdRequired & (b_AnyModuleRequired = FALSE) then
          b_AnyModuleRequired := TRUE;
          // if any access is required => the businterface is also required
          tempCmd.uiCmd := _BUS_IF_SET_REQUIRED;
          ToBusInterface.NewInst(pPara:=#tempCmd, pResult:=#_result);
          if _result.aData[0]$t_BusIFRetvalErrorcode <> _BUS_IF_RETVAL_OK then
            LogError("@03DE (SdiasSafetyManagerFSoE::HGWOut::NewInst) Failed to set the BusInterface to required");
          end_if;
        end_if;
      else
          ret_code := ERROR;
        end_if;

      else
        // unknown version of the request
        ret_code := ERROR;
      end_if;

    //**********************************************************************************************************************************************************
    CMD_SM_ADD_ROUTING_INFO:
      tempHWPath.p_us_Path := NIL;
      tempHWPath.p_us_PathComp := NIL;
      tempHWPath.ui_PathCompLen := 0;
      if sHGW.hdSafetyNrb <> pPara^.aPara[0]$HDINT then
        //safe act hgw safety number
        sHGW.hdSafetyNrb := pPara^.aPara[0]$HDINT;
        //add routing element for hgw panel
        dRetCode := AddRoutingElement(ud_SafeNumber:=sHGW.hdSafetyNrb, ud_thisp:=sHGW.pThis$UDINT, pObject:=#tempHWPath);
        if dRetCode <> 0 then
          ret_code := ERROR;
        end_if;
      end_if;

    //**********************************************************************************************************************************************************
    CMD_SM_ADD_SDO_TO_BUFFER:
      ret_code := ClassSvr.NewInst(pPara:=pPara, pResult:=pResult);

  //**********************************************************************************************************************************************************

  else
    //if command is not known send it to safety manager
    if pSafetyManagerThis then
      ret_code := pSafetyManagerThis^.NewInst(pPara, pResult);
    end_if;

  end_case;

END_FUNCTION

FUNCTION VIRTUAL SdiasSafetyManagerFSoE::SafeActModuleConfig
  VAR_INPUT
    sActModuleConfig 	: t_ModuleCfg;
  END_VAR

  sCPUConfig := sActModuleConfig;

END_FUNCTION

FUNCTION VIRTUAL GLOBAL SdiasSafetyManagerFSoE::FCN_Command::Write
  VAR_INPUT
    input (EAX) 	: UDINT;
  END_VAR
  VAR_OUTPUT
    result (EAX) 	: UDINT;
  END_VAR

  // only if input is valid and we're in the right state
  if (input = 1) & (FCN_StateMachine = 1) then
    sFlexCon.CommandRequest := input;
  end_if;

  result := input;

END_FUNCTION
